(* IEC 61131-3 sources: volt/packages/volt-lsp-iec/test-corpus/pro2193/Device/Plc Logic/Application/09 Misc, 2 files *)

(* ---- eExceptionCodes.dut ---- *)
{attribute 'qualified_only'}
{attribute 'strict'}
TYPE eExceptionCodes :
(
	DashboardTask := 0,
	EdgePcTask,
	Ethernet,
	JsonTask,
	MainTask,
	RecipeTask,
	InjectionMouldingMachine,
	LabelSuppliers,
	CassetteAdjustment,
	Magazines,
	XiUnits,
	XuUnits,
	YUnits,
	RejectStations,
	Chains,
	ZUnits,
	ZRUnits,
	VisionSystems,
	Conveyors,
	Fanucs,
	BufferRacks,
	BoxInfeeds,
	BoxCenterUnits,
	BoxPushers,
	BoxOutfeeds,
	TimeSettings,
	EtherCAT_Diag,
	ErrorHandling,
	HardwareButtons,
	BfuButtons,
	HMI,
	HMI_BFU,
	HardwareUnits,
	ProcessModules,
	SER,
	BFU,
	IQ_Handling
);
END_TYPE

(* ---- GVL_Exceptions.gvl ---- *)
{attribute 'qualified_only'}
VAR_GLOBAL
	xException : BOOL;
	aeExceptionCodes: ARRAY[0..50] OF __SYSTEM.ExceptionCode;
	iCounter	: UDINT;
END_VAR
